{attribute 'qualified_only'}
{attribute 'strict'}
{attribute 'to_string'}
TYPE E_OpMode : (
		manual := 0,
		auto
	);
END_TYPE

(* stored: Version 1.1.0.1
   DUT E_OpMode: Id {8443ccac-7148-4542-8a1d-551519071d8c} *)
